ABB RAPID module: CalibData.modx

MODULE CalibData
    PERS tooldata MyTool:=[TRUE,[[31.792631019,-0,229.638935148],[0.945518576,0,0.325568154,0]],[1,[0,0,1],[1,0,0,0],0,0,0]];
    PERS wobjdata Koordinatensystem_Modul5:=[FALSE,TRUE,"",[[-499.960321416,1020.013088225,257.5],[1,0,0,0.000005866]],[[0,0,0],[1,0,0,0]]];
    PERS wobjdata Koordinatensystem_Modul2:=[FALSE,TRUE,"",[[498.985385611,-1020.52304872,257.5],[0.000473151,0,0,-0.999999888]],[[0,0,0],[1,0,0,0]]];
    PERS wobjdata Koordinatensystem_Modul1:=[FALSE,TRUE,"",[[1134.907540478,-83.031342842,257.5],[0.500647833,0,0,-0.865651054]],[[0,0,0],[1,0,0,0]]];
    PERS wobjdata Koordinatensystem_Modul3:=[FALSE,TRUE,"",[[-636.650058157,-941.997300822,257.5],[0.50036151,0,0,0.865816585]],[[0,0,0],[1,0,0,0]]];
    PERS wobjdata Koordinatensystem_Modul4:=[FALSE,TRUE,"",[[-1133.976818569,78.784535634,257.5],[0.86565239,0,0,0.500645524]],[[0,0,0],[1,0,0,0]]];
    PERS wobjdata Koordinatensystem_Modul6:=[FALSE,TRUE,"",[[638.159114859,940.449669808,257.5],[0.866179246,-0,0,-0.499733442]],[[0,0,0],[1,0,0,0]]];
    PERS wobjdata coordinate_system_module_5:=[FALSE,TRUE,"",[[-499.960321416,1020.013088225,257.5],[1,0,0,0.000005866]],[[0,0,0],[1,0,0,0]]];
    PERS wobjdata coordinate_system_module_2:=[FALSE,TRUE,"",[[498.985385611,-1020.52304872,257.5],[0.000473151,0,0,-0.999999888]],[[0,0,0],[1,0,0,0]]];
    PERS wobjdata coordinate_system_module_1:=[FALSE,TRUE,"",[[1134.907540478,-83.031342842,257.5],[0.500647833,0,0,-0.865651054]],[[0,0,0],[1,0,0,0]]];
    PERS wobjdata coordinate_system_module_3:=[FALSE,TRUE,"",[[-636.650058157,-941.997300822,257.5],[0.50036151,0,0,0.865816585]],[[0,0,0],[1,0,0,0]]];
    PERS wobjdata coordinate_system_module_4:=[FALSE,TRUE,"",[[-1133.976818569,78.784535634,257.5],[0.86565239,0,0,0.500645524]],[[0,0,0],[1,0,0,0]]];
    PERS wobjdata coordinate_system_module_6:=[FALSE,TRUE,"",[[638.159114859,940.449669808,257.5],[0.866179246,-0,0,-0.499733442]],[[0,0,0],[1,0,0,0]]];
ENDMODULE
